DATA_BLOCK "db3100_BC400_Chaves"
TITLE = db3100_BC400_Chaves v0.2 (DB3100)
{ S7_Optimized_Access := 'FALSE' }
AUTHOR : 'Reginaldo Lobo'
VERSION : 0.2
NON_RETAIN
////====================================
//// db3100_BC400_Chaves (DB3100) - GERADO por plc/bt2/gerador/gerar_banco_v0.2.py (03/11/2026) - nao compilado no TIA, nao testado
//// O QUE FAZ : mesmo papel do db150_BC56_Chaves v0.3, arrays de 16 chaves. Banco BC400: 13 chaves reais, 3 reserva. FB: FB100/FB101.
//// OFFSETS (calculados; CONFERIR na coluna "Deslocamento" do TIA): cb.ligar X0.0 | sb.ligada X2.0 | habilitada X4.0 | setupOk X6.0
////    kwReal D8 | rMedidoOhm D72 | rTeoricoOhm D136 | setupData B200 (12 bytes cada) | nominal D392
////    chaveSel W456 | salvar X458.0 | usarKwReal X458.1 | cbBanco.ligar X460.0 | sbBanco.seletoraAuto X462.0 | comEt200Ok X462.1
//// kW nominal na ordem fisica das chaves (informado pelo operador em 30/10/2026).
////=====================================
   VAR
      cb : Struct
         ligar : Array[1..16] of Bool;
      END_STRUCT;

      sb : Struct
         ligada : Array[1..16] of Bool;
      END_STRUCT;

      setup : Struct
         habilitada   : Array[1..16] of Bool;
         setupOk      : Array[1..16] of Bool;
         kwReal       : Array[1..16] of Real;
         rMedidoOhm   : Array[1..16] of Real;
         rTeoricoOhm  : Array[1..16] of Real;
         setupData    : Array[1..16] of DTL;
         nominal      : Array[1..16] of Real;
         chaveSel     : UInt;
         salvar       : Bool;
         usarKwReal   : Bool;
      END_STRUCT;

      cbBanco : Struct   // DBX460.0
         ligar : Bool;
      END_STRUCT;

      sbBanco : Struct   // DBX462.0
         seletoraAuto : Bool;
         comEt200Ok : Bool;
      END_STRUCT;
   END_VAR


BEGIN
   setup.nominal[1] := 5.0;
   setup.nominal[2] := 5.0;
   setup.nominal[3] := 10.0;
   setup.nominal[4] := 10.0;
   setup.nominal[5] := 10.0;
   setup.nominal[6] := 10.0;
   setup.nominal[7] := 50.0;
   setup.nominal[8] := 50.0;
   setup.nominal[9] := 50.0;
   setup.nominal[10] := 50.0;
   setup.nominal[11] := 50.0;
   setup.nominal[12] := 50.0;
   setup.nominal[13] := 50.0;
   // 14..16: reserva, 0.0

END_DATA_BLOCK
